//---------------------------------------------------------------------------------------------------------------
//
//  HAUD 2026.10.20
//
//
//  fb_DistributorByTicket
//  - uses 1 XtsStation via _ItfProcessCollector
//  - this instance checks its process list for an entry (Count > 0)
//      - pops ticket data from top of the list (GetHead)
//      - sends the mover to target stations according to bitmask in ST_PROCESS_DATA.wTarget
//
//  - inherits fb_Instance, which provides a design pattern in order to build different specific processes in a structured way
//  - used for targeting movers to predetermined bitmask of substations (one to many)
//
//
//  - constructed with fb_Instance main state (_eState) in addition to a substate (_eStateProgress)
//  - substate enables to handle procedures within main state by preventing race conditions 
//    with the help of small steps and decisions with clear separation from each other 
//
//---------------------------------------------------------------------------------------------------------------//
// This SOFTWARE is provided as an Exemple by THE PROVIDER "as is" and "with all faults." THE PROVIDER makes no  //
// representations or warranties of any kind concerning the safety, suitability, lack of viruses, inaccuracies,  //
// typographical errors, or other harmful components of this SOFTWARE. There are inherent dangers in the use of  //
// any software, and you are solely responsible for determining whether this SOFTWARE is compatible with your    //
// equipment and other software installed on your equipment. You are also solely responsible for the protection  //
// of your equipment and backup of your data, and THE PROVIDER will not be liable for any damages you may suffer //
// in connection with using, modifying, or distributing this SOFTWARE.                                           //
//---------------------------------------------------------------------------------------------------------------//
FUNCTION_BLOCK fb_DistributorByTicket EXTENDS fb_Instance
VAR
  //----------------------------------------------------------------------------------
  // outfeed target must be initialized with a valid target
  // I just use the default target that I am going to use in the basic process setup
  // this target is then updated and checked on arrival of a process ticket
  //----------------------------------------------------------------------------------
  _nProcessTarget               : E_INSTANCE;     // to whom am I connected --> to the data from the ticket
  //----------------------------------------------------------------------------------

  // target XTS station range
  _nTargetStationLast           : UINT;           // where does the target process end
  _nTargetStationFirst          : UINT;           // where does the target process start

  _WriteResult                  : ST_PROCESS_LIST_RESULT;   // last job written to target
  _DeleteResult                 : ST_PROCESS_LIST_RESULT;   // last job executed

  _nPrc                         : E_INSTANCE;
  _nTarget                      : E_INSTANCE;

  _idx                          : UINT;
  _nTargetIndex                 : ARRAY[1..SIZEOF(T_PROCESS)*8] OF USINT;

  _MoverInfo                    : ST_MOVER_INFO;      // Information from the Mover in Station
  _StationState                 : ST_STATION_STATE;   // BufferInfeed has only one XtsStation to work
END_VAR

//-----------------------------------------------------------------------------
//-----------------------------------------------------------------------------
// check pointer and interface
// connect Ctrl/State to _ItfProcessCollector
// set message device identification
//-----------------------------------------------------------------------------
IF NOT Check() THEN 
  RETURN; 
END_IF
//-----------------------------------------------------------------------------
// check command
//-----------------------------------------------------------------------------
_eCmd                                         := _stInstanceCtrl[_nProcess].Cmd;
IF (_eCmd <> _eCmdOld)
THEN
  CASE _eCmd
  OF
    E_INSTANCE_CMD.INIT:
      // clear init info
      _eInit                                  := _ItfProcessCollector[_nProcess].Init(FALSE);
  
      IF _ItfProcessList[_nProcess].InitList()  // clear linked list
      THEN
        Clear();
        _eStateInstance                       := E_INSTANCE_STATE.INIT;
        _eStateProgress                       := E_PROGRESS.PROGRESS_INIT;
      END_IF
  END_CASE
  CmdLog();
  _eCmdOld                                    := _eCmd;
END_IF
//-----------------------------------------------------------------------------
// cyclic information of mover and station
//-----------------------------------------------------------------------------
_StationState                                 := _ItfProcessCollector[_nProcess].GetStationState  (_ItfProcessCollector[_nProcess].StationLast);
//-----------------------------------------------------------------------------
//-----------------------------------------------------------------------------
// state machine for BufferInfeed work
//-----------------------------------------------------------------------------
CASE _eStateInstance
OF
  E_INSTANCE_STATE.NULL:
    // first cycle startup
    // initialize linked list, clears all entries
    IF _ItfProcessList[_nProcess].InitList()
    THEN
      _eInit                                  := _ItfProcessCollector[_nProcess].Init(FALSE);
      _eStateProgress                         := E_PROGRESS.PROGRESS_INIT;
      _eStateInstance                         := E_INSTANCE_STATE.INIT;
    END_IF


  E_INSTANCE_STATE.INIT:
    //-------------------------------------------------------------------------
    CASE _eStateProgress
    OF
    // E_INSTANCE_STATE.INIT:
    //-------------------------------------------------------------------------
      E_PROGRESS.PROGRESS_ERROR:
        IF (_nProcessTarget > 0) AND
           (_nProcessTarget < E_INSTANCE.INSTANCE_MAX)
        THEN
          _eStateProgress                     := E_PROGRESS.PROGRESS_INIT;
        END_IF

    // E_INSTANCE_STATE.INIT:
    //-------------------------------------------------------------------------
      E_PROGRESS.PROGRESS_INIT:
        IF NOT (_nProcessTarget > 0) OR
           NOT (_nProcessTarget < E_INSTANCE.INSTANCE_MAX)
        THEN
          _eStateProgress                     := E_PROGRESS.PROGRESS_ERROR;

        ELSE
          _eStateProgress                     := E_PROGRESS.PROGRESS_BUSY;
        END_IF

    // E_INSTANCE_STATE.INIT:
    //-------------------------------------------------------------------------
      E_PROGRESS.PROGRESS_BUSY:
        // wait for process collector check to be done
        //  - checks range of XtsStations
        //  - checks count of XtsStations
        IF (_stCollectorState.Check = E_PROCESS_CHECK.CHECK_DONE)
        THEN
          _eInit                              := _ItfProcessCollector[_nProcess].Init(TRUE);
  
          IF (_eInit = E_PROGRESS.PROGRESS_DONE)
          THEN
            IF NOT (_nProcessTarget > 0) OR
               NOT (_nProcessTarget < E_INSTANCE.INSTANCE_MAX)
            THEN
              // an invalid target you must have not
              _eStateProgress                 := E_PROGRESS.PROGRESS_ERROR;

              _stMsg.eType                    := E_MessageType.eMessageError;
              _stMsg.eSubdevice               := e_Subdevice.Instance_DistributorByTicket;
              _stMsg.iErrorNumber             := _nProcessTarget;
              _stMsg.sText                    := concat(TO_STRING(_eStateInstance), ': ProcessTarget: ');
              _stMsg.sText                    := concat(_stMsg.sText, TO_STRING(_eStateProgress));
              f_MessageSet(_stMsg);

            ELSE
              _ItfProcessCollector[_nProcess].Init(FALSE); // clear init procedure

              // initialization of BufferInfeed: _ItfProcessCollector with XtsStation
              _stCollectorCtrl.Cmd            := E_PROCESS_CTRL.PROCESS_DISABLE;  // switch off _ItfProcessCollector and XtsStation
              _eStateProgress                 := E_PROGRESS.PROGRESS_INIT;        // clear sub state
              _eStateInstance                 := E_INSTANCE_STATE.DISABLED;       // switch to disabled as default after startup
            END_IF
          END_IF
        END_IF
    END_CASE
END_CASE
//-----------------------------------------------------------------------------
// DISABLED:
//  - clear local list result data
//  - wait for enable from the outside
//-----------------------------------------------------------------------------
CASE _eStateInstance
OF
  E_INSTANCE_STATE.DISABLED:
    //-------------------------------------------------------------------------
    CASE _eStateProgress
    OF
      E_PROGRESS.PROGRESS_INIT:
        _stCollectorCtrl.Cmd                  := E_PROCESS_CTRL.PROCESS_DISABLE;  // switch off _ItfProcessCollector and XtsStation
        _eStateProgress                       := E_PROGRESS.PROGRESS_BUSY;
        // clear data for a new round
        memset(ADR(_stListResult), 0, SIZEOF(_stListResult));

        _stCollectorCtrl.ActivateStation      := 0; // clear activation mask of my process
        _stCollectorCtrl.NestMask             := 1; // my process target has one nest

        _nPrc                                 := _nProcess;
        _nTarget                              := _nProcessTarget;
    END_CASE
    // E_INSTANCE_STATE.DISABLED:
    //-------------------------------------------------------------------------
    CASE _eStateProgress
    OF
      E_PROGRESS.PROGRESS_BUSY:
        CASE _eCmd
        OF
          E_INSTANCE_CMD.ENABLE:              // turn it on!!
            _nPrc                             := _nProcess;
            _nTarget                          := _nProcessTarget;

            _eStateInstance                   := E_INSTANCE_STATE.DETECTION;
            _eStateProgress                   := E_PROGRESS.PROGRESS_BUSY;
  
            IF (_MessageLevel > E_MessageType.eMessageInfo)
            THEN
              _stMsg.eType                    := E_MessageType.eMessageVerbose;
              _stMsg.eSubdevice               := e_Subdevice.Instance_DistributorByTicket;
              _stMsg.iErrorNumber             := 0;
              _stMsg.sText                    := concat(TO_STRING(_eStateInstance), ': ');
              _stMsg.sText                    := concat(_stMsg.sText, TO_STRING(_eStateProgress));
              f_MessageSet(_stMsg);
            END_IF

        END_CASE
    END_CASE
END_CASE
//-----------------------------------------------------------------------------
// DETECTION: 
//  - check inked list and GetHead()
//  - copy job data
//  - switch on process
//-----------------------------------------------------------------------------
CASE _eStateInstance
OF
  E_INSTANCE_STATE.DETECTION:
    //-------------------------------------------------------------------------
    CASE _eStateProgress
    OF
      E_PROGRESS.PROGRESS_BUSY:
        IF (_eCmd = E_INSTANCE_CMD.DISABLE)
        THEN
          _eStateInstance                     := E_INSTANCE_STATE.DISABLED;
          _eStateProgress                     := E_PROGRESS.PROGRESS_INIT;

        ELSIF (_ItfProcessList[_nPrc].Count > 0)
        THEN
          // get new job order for my process
          // check my list for a new round of movers
          _stListResult                       := _ItfProcessList[_nPrc].GetHead();  // the list results carries information about the requirements of the target process (who and where)

          IF (_stListResult.wState <> 0)
          THEN
            // error in list results must not appear
            // if you land here, there is somethng wrong with the initialization or configuration of the linked list
            _eStateProgress                   := E_PROGRESS.PROGRESS_ERROR;

            _stMsg.eType                      := E_MessageType.eMessageError;
            _stMsg.eSubdevice                 := e_Subdevice.Process_LinkedList_GetHead;
            _stMsg.iErrorNumber               := _stListResult.wState;
            _stMsg.sText                      := concat(TO_STRING(_eStateInstance), ': _ListResult.wState: ');
            _stMsg.sText                      := concat(_stMsg.sText, TO_STRING(_eStateProgress));
            f_MessageSet(_stMsg);

          ELSE
            IF (_MessageLevel > E_MessageType.eMessageError)
            THEN
              _stMsg.eType                    := E_MessageType.eMessageInfo;
              _stMsg.eSubdevice               := e_Subdevice.Process_LinkedList_GetHead;
              _stMsg.iErrorNumber             := _nPrc;
              _stMsg.sText                    := concat(TO_STRING(_eStateInstance), ': ');
              _stMsg.sText                    := concat(_stMsg.sText, '_ListResult.stData.wTarget: ');
              _stMsg.sText                    := concat(_stMsg.sText, _ItfProcessCollector[_nPrc].BitsToString(_stListResult.stData.wTarget));
              f_MessageSet(_stMsg);
            END_IF

            _stProcessData                    := _stListResult.stData;  // list result contains data for target process

            IF (_stProcessData.wTarget > 0)
            THEN
              _eStateProgress                 := E_PROGRESS.PROGRESS_CHECK;

              IF (_MessageLevel = E_MessageType.eMessageBatch)
              THEN
                _stMsg.eType                  := E_MessageType.eMessageBatch;
                _stMsg.eSubdevice             := e_Subdevice.Instance_DistributorByTicket;
                _stMsg.iErrorNumber           := _nPrc;
                _stMsg.sText                  := concat(TO_STRING(_eStateProgress), ': ');
                _stMsg.sText                  := concat(_stMsg.sText, TO_STRING(e_message_batch.MSG_BATCH_JOB_STARTED));
                f_MessageSet(_stMsg);
              END_IF
            ELSE
              _DeleteResult                   := _ItfProcessList[_nPrc].RemoveHeadValue();
            END_IF

            // check target mask for entries
            IF NOT (_stProcessData.wTarget > 0)
            THEN
              _stMsg.eType                    := E_MessageType.eMessageWarning;
              _stMsg.eSubdevice               := e_Subdevice.Instance_DistributorByTicket;
              _stMsg.iErrorNumber             := 666;
              _stMsg.sText                    := concat(TO_STRING(_eStateInstance), ': ');
              _stMsg.sText                    := concat(_stMsg.sText, '_ProcessData.wTarget: ');
              _stMsg.sText                    := concat(_stMsg.sText, _ItfProcessCollector[_nProcess].BitsToString(_stProcessData.wTarget));
              f_MessageSet(_stMsg);
            END_IF
          END_IF
        END_IF
    END_CASE
    // E_INSTANCE_STATE.DETECTION
    //-------------------------------------------------------------------------
    CASE _eStateProgress
    OF
      E_PROGRESS.PROGRESS_CHECK:
        // do some plausibility checks on the ticket data
        IF NOT (_stProcessData.nTargetId > 0) OR
           NOT (_stProcessData.nTargetId < E_INSTANCE.INSTANCE_MAX) OR
           NOT (_stProcessData.nTargetId <> _nProcess)
        THEN
          _stMsg.eType                        := E_MessageType.eMessageError;
          _stMsg.eSubdevice                   := e_Subdevice.Instance_DistributorByTicket;
          _stMsg.iErrorNumber                 := _stProcessData.nTargetId;
          _stMsg.sText                        := concat(TO_STRING(_eStateInstance), ': _stProcessData.nTargetId: ');
          _stMsg.sText                        := concat(_stMsg.sText, TO_STRING(E_PROGRESS.PROGRESS_ERROR));
          f_MessageSet(_stMsg);

          // not a plausible target, delete ticket and go back to checking the list
          _DeleteResult                       := _ItfProcessList[_nPrc].RemoveHeadValue();
          _eStateProgress                     := E_PROGRESS.PROGRESS_BUSY;
        ELSE
          // update target data with ticket data
          _nTarget                            := _stProcessData.nTargetId;
          _nTargetStationLast                 := _ItfProcessCollector[_nTarget].StationLast;
          _nTargetStationFirst                := _ItfProcessCollector[_nTarget].StationFirst;

          IF (_ItfProcessCollector[_nTarget].ProcessState.Check = E_PROCESS_CHECK.CHECK_DONE)
          THEN
            _eStateProgress                   := E_PROGRESS.PROGRESS_WORKING;

            IF (_MessageLevel > E_MessageType.eMessageWarning)
            THEN
              _stMsg.eType                    := E_MessageType.eMessageInfo;
              _stMsg.eSubdevice               := e_Subdevice.Instance_DistributorByTicket;
              _stMsg.iErrorNumber             := _stProcessData.nTargetId;
              _stMsg.sText                    := concat(TO_STRING(_stProcessData.nProcessId), ': _stProcessData.nTargetId: ');
              _stMsg.sText                    := concat(_stMsg.sText, TO_STRING(_eStateProgress));
              f_MessageSet(_stMsg);
            END_IF
          END_IF
        END_IF
    END_CASE
    // E_INSTANCE_STATE.DETECTION
    //-------------------------------------------------------------------------
    CASE _eStateProgress
    OF
      E_PROGRESS.PROGRESS_WORKING:
        // check for disabled process interface state
        CASE _stCollectorState.State
        OF
          E_PROCESS_STATE.PROCESS_DISABLE:

          CASE _stCollectorState.Result
          OF
            E_PROGRESS.PROGRESS_BUSY:         // busy from _State.Result means, waiting for input
              // now the preparation for the target process may begin
              _stCollectorCtrl.Cmd               := E_PROCESS_CTRL.PROCESS_ENABLE; // switch on my state machine in _ItfProcessCollector
              _stCollectorCtrl.ActivateStation   := 1;                             // enable my XtsStation in _ItfProcessCollector (BufferInfeed has only one XtsStation)

              _eStateInstance                 := E_INSTANCE_STATE.ENABLED;         // go check if my process is switched on
              _eStateProgress                 := E_PROGRESS.PROGRESS_INIT;         // reset substate

              IF (_MessageLevel > E_MessageType.eMessageInfo)
              THEN
                _stMsg.eType                  := E_MessageType.eMessageVerbose;
                _stMsg.eSubdevice             := e_Subdevice.Instance_DistributorByTicket;
                _stMsg.iErrorNumber           := 0;
                _stMsg.sText                  := concat(TO_STRING(_eStateInstance), ': ');
                _stMsg.sText                  := concat(_stMsg.sText, TO_STRING(_eStateProgress));
                f_MessageSet(_stMsg);
              END_IF
          END_CASE
        END_CASE
    END_CASE
END_CASE
//-----------------------------------------------------------------------------
// ENABLED
//  - check process for enabled stations from list entry
//  - switch to sending
//  - allow movers to be sent
//-----------------------------------------------------------------------------
CASE _eStateInstance
OF
  E_INSTANCE_STATE.ENABLED:
    //-------------------------------------------------------------------------
    CASE _eStateProgress
    OF
      E_PROGRESS.PROGRESS_INIT:
        CASE _stCollectorState.State
        OF
          E_PROCESS_STATE.PROCESS_ENABLE:
          CASE _stCollectorState.Result
          OF
            E_PROGRESS.PROGRESS_BUSY:
              // now my process and all XtsStations within are switched on
              // check infeed into my process
              _stCollectorCtrl.Cmd            := E_PROCESS_CTRL.PROCESS_STATIONS_SEND; // tells my process to go check the infeed
              _eStateProgress                 := E_PROGRESS.PROGRESS_BUSY; // go check how the infeed into my process is doing

              IF (_MessageLevel > E_MessageType.eMessageWarning)
              THEN
                _stMsg.eType                  := E_MessageType.eMessageInfo;
                _stMsg.eSubdevice             := e_Subdevice.Instance_DistributorByTicket;
                _stMsg.iErrorNumber           := _StationState.nMoverId;
                _stMsg.sText                  := concat(TO_STRING(_eStateInstance), ': ');
                _stMsg.sText                  := concat(_stMsg.sText, TO_STRING(_eStateProgress));
                f_MessageSet(_stMsg);
              END_IF
          END_CASE
        END_CASE
    END_CASE
    // E_INSTANCE_STATE.ENABLED:
    //-------------------------------------------------------------------------
    CASE _eStateProgress
    OF
      E_PROGRESS.PROGRESS_BUSY:
        CASE _stCollectorState.State
        OF
          E_PROCESS_STATE.PROCESS_STATIONS_OUTFEED:
          CASE _stCollectorState.Result       // if collector is ready to send mover
          OF
            E_PROGRESS.PROGRESS_BUSY:
              // check if the mover is in range
              IF (_rCheckPositionEnd > _rCheckPositionStart)
              THEN
                IF (_StationState.rMoverModPos > _rCheckPositionStart) AND
                   (_StationState.rMoverModPos < _rCheckPositionEnd)
                THEN
                  _eStateProgress             := E_PROGRESS.PROGRESS_PREPARE;
                END_IF
              ELSE
                IF (_StationState.rMoverModPos > _rCheckPositionStart) OR
                   (_StationState.rMoverModPos < _rCheckPositionEnd)
                THEN
                  _eStateProgress             := E_PROGRESS.PROGRESS_PREPARE;
                END_IF
              END_IF
          END_CASE
        END_CASE
    END_CASE
    // E_INSTANCE_STATE.ENABLED:
    //-------------------------------------------------------------------------
    CASE _eStateProgress
    OF
      E_PROGRESS.PROGRESS_PREPARE:
        // now we know the mover is in range
        // continue to finish
        _stCollectorCtrl.Cmd                  := E_PROCESS_CTRL.PROCESS_STATIONS_SEND;

        _eStateInstance                       := E_INSTANCE_STATE.FINISH;   // go get data ready for outfeed
        _eStateProgress                       := E_PROGRESS.PROGRESS_INIT;  // reset substate

        IF (_MessageLevel > E_MessageType.eMessageError)
        THEN
          _stMsg.eType                        := E_MessageType.eMessageInfo;
          _stMsg.eSubdevice                   := e_Subdevice.Instance_DistributorByTicket;
          _stMsg.iErrorNumber                 := _StationState.nMoverId;
          _stMsg.sText                        := concat(TO_STRING(_eStateInstance), ': ');
          _stMsg.sText                        := concat(_stMsg.sText, TO_STRING(_eStateProgress));
          f_MessageSet(_stMsg);
        END_IF
    END_CASE
END_CASE
//-----------------------------------------------------------------------------
// FINISH:
//  - write target (Last to First)
//  - delete target bit from linked list result (_ProcessData.wTarget)
//  - send out mover
//  - check _ProcessData.wTarget for next mover
//  - check if all movers in job were sent (ProcessData.wTarget = 0)
//  - RemoveHead() from my list
//  - AddTail() at TargetProcess
//  - check to proceed
//-----------------------------------------------------------------------------
CASE _eStateInstance
OF
  E_INSTANCE_STATE.FINISH:
    //-------------------------------------------------------------------------
    CASE _eStateProgress
    OF
      E_PROGRESS.PROGRESS_INIT:
      // check bit mask for sending mover to required targets
      // get target index for mover from process list entry
      FOR _idx := _nTargetStationLast TO _nTargetStationFirst BY(-1)
      DO
        IF (ItfProcessCollector[_nPrc].BitGet(_stProcessData.wTarget, _idx-_nTargetStationFirst))
        THEN
          _eStateProgress                     := E_PROGRESS.PROGRESS_BUSY;

          _nTargetIndex[1]                    := TO_USINT(_idx);
          _ItfProcessCollector[_nPrc].TargetIndex := _nTargetIndex; // write Xts target onto my ProcessCollector interface

          // got the target, now delete the just found bit of this job
          _stProcessData.wTarget              := _ItfProcessCollector[_nPrc].
                                                 BitDel(_stProcessData.wTarget, _idx-_nTargetStationFirst);

          IF (_MessageLevel > E_MessageType.eMessageVerbose)
          THEN
            _stMsg.eType                      := E_MessageType.eMessageSentient;
            _stMsg.eSubdevice                 := e_Subdevice.Instance_DistributorByTicket;
            _stMsg.iErrorNumber               := _idx;
            _stMsg.sText                      := concat('_ProcessData.wTarget: ', 
                                                 _ItfProcessCollector[_nPrc].BitsToString(_stProcessData.wTarget));
            f_MessageSet(_stMsg);
          END_IF
          EXIT;
        END_IF
      END_FOR
    END_CASE
    // E_INSTANCE_STATE.FINISH:
    //-------------------------------------------------------------------------
    CASE _eStateProgress
    OF
      E_PROGRESS.PROGRESS_BUSY:
        CASE _stCollectorState.State
        OF
          E_PROCESS_STATE.PROCESS_STATIONS_OUTFEED: // double check my process' state
          CASE _stCollectorState.Result
          OF
            E_PROGRESS.PROGRESS_BUSY:
              // now data is prepared and copied to the right places
              _stCollectorCtrl.Cmd            := E_PROCESS_CTRL.PROCESS_STATIONS_OUTFEED; // tell my process to release the mover
              _eStateProgress                 := E_PROGRESS.PROGRESS_CHECK; // go check for more to do

              IF (_MessageLevel > E_MessageType.eMessageInfo)
              THEN
                _stMsg.eType                  := E_MessageType.eMessageVerbose;
                _stMsg.eSubdevice             := e_Subdevice.Instance_DistributorByTicket;
                _stMsg.iErrorNumber           := _nPrc;
                _stMsg.sText                  := concat(TO_STRING(_eStateInstance), ': ');
                _stMsg.sText                  := concat(_stMsg.sText, TO_STRING(_eStateProgress));
                f_MessageSet(_stMsg);
              END_IF
          END_CASE
        END_CASE
    END_CASE
    // E_INSTANCE_STATE.FINISH:
    //-------------------------------------------------------------------------
    CASE _eStateProgress
    OF
      E_PROGRESS.PROGRESS_CHECK:
        CASE _stCollectorState.State
        OF
          E_PROCESS_STATE.PROCESS_DISABLE:
            IF (_stProcessData.wTarget <> 0)
            THEN
              _stCollectorCtrl.Cmd               := E_PROCESS_CTRL.PROCESS_ENABLE; // switch on my state machine in _ItfProcessCollector
              _stCollectorCtrl.ActivateStation   := 1;                             // enable my XtsStation in _ItfProcessCollector (BufferInfeed has only one XtsStation)

              _eStateInstance                 := E_INSTANCE_STATE.ENABLED;         // go check if my process is switched on
              _eStateProgress                 := E_PROGRESS.PROGRESS_INIT;         // reset substate

              IF (_MessageLevel > E_MessageType.eMessageInfo)
              THEN
                _stMsg.eType                  := E_MessageType.eMessageVerbose;
                _stMsg.eSubdevice             := e_Subdevice.Instance_DistributorByTicket;
                _stMsg.iErrorNumber           := _nPrc;
                _stMsg.sText                  := concat(TO_STRING(_eStateInstance), ': ');
                _stMsg.sText                  := concat(_stMsg.sText, TO_STRING(_eStateProgress));
                f_MessageSet(_stMsg);
              END_IF
            ELSE
              // job done, all movers were sent
              // job done, delete from top of my list
              _DeleteResult                   := _ItfProcessList[_nPrc].RemoveHeadValue();

              IF (_DeleteResult.wState <> 0)
              THEN
                // deleting from list must be successful
                // IF you land here, there is something wrong with initialization or configuration of the linked list
                _eStateProgress               := E_PROGRESS.PROGRESS_ERROR;
              ELSE
                _eStateProgress               := E_PROGRESS.PROGRESS_WORKING; // job is done, now go and write ticket to _nTargetProcess
              END_IF
            END_IF 
        END_CASE
    END_CASE
    // E_INSTANCE_STATE.FINISH:
    //-------------------------------------------------------------------------
    CASE _eStateProgress
    OF
      E_PROGRESS.PROGRESS_WORKING:
        // write process ticket, then go back up
        //_WriteResult                          := _ItfProcessList[_nTarget].AddTailValue(_stListResult.stData);

        IF (_WriteResult.wState <> 0)
        THEN
          // adding to target list must be successful on the first try
          // IF you land here, there is something wrong with initialization or configuration of the linked list
          _eStateProgress                     := E_PROGRESS.PROGRESS_ERROR;
        ELSE
          _eStateProgress                     := E_PROGRESS.PROGRESS_DONE;

          IF (_MessageLevel > E_MessageType.eMessageError)
          THEN
            _stMsg.eType                      := E_MessageType.eMessageInfo;
            _stMsg.eSubdevice                 := e_Subdevice.Process_LinkedList_AddTail;
            _stMsg.iErrorNumber               := _nTarget;
            _stMsg.sText                      := concat(TO_STRING(_eStateInstance), ': ');
            _stMsg.sText                      := concat(_stMsg.sText, TO_STRING(_eStateProgress));
            //f_MessageSet(_stMsg);
          END_IF
          IF (_MessageLevel = E_MessageType.eMessageBatch)
          THEN
            _stMsg.eType                      := E_MessageType.eMessageBatch;
            _stMsg.eSubdevice                 := e_Subdevice.Instance_DistributorByTicket;
            _stMsg.iErrorNumber               := _nPrc;
            _stMsg.sText                      := concat(TO_STRING(_eStateProgress), ': ');
            _stMsg.sText                      := concat(_stMsg.sText, TO_STRING(e_message_batch.MSG_BATCH_JOB_DONE));
            f_MessageSet(_stMsg);
          END_IF
        END_IF
    END_CASE
    // E_INSTANCE_STATE.FINISH:
    //-------------------------------------------------------------------------
    CASE _eStateProgress
    OF
      E_PROGRESS.PROGRESS_DONE:
        //----------------------------------
        //  wait for command from higher up
        //----------------------------------
        CASE _eCmd
        OF
          // command to disable required
          E_INSTANCE_CMD.DISABLE:
            _eStateInstance                   := E_INSTANCE_STATE.DISABLED;
            _eStateProgress                   := E_PROGRESS.PROGRESS_INIT;

            IF (_MessageLevel > E_MessageType.eMessageInfo)
            THEN
              _stMsg.eType                    := E_MessageType.eMessageVerbose;
              _stMsg.eSubdevice               := e_Subdevice.Instance_DistributorByTicket;
              _stMsg.iErrorNumber             := _nPrc;
              _stMsg.sText                    := concat(TO_STRING(_eStateInstance), ': ');
              _stMsg.sText                    := concat(_stMsg.sText, TO_STRING(_eStateProgress));
              f_MessageSet(_stMsg);
            END_IF
        END_CASE
    END_CASE
END_CASE
//-----------------------------------------------------------------------------
//-----------------------------------------------------------------------------
_stInstanceState[_nProcess].ProcessIdentity   := _nProcess;
_stInstanceState[_nProcess].ProcessState      := _eStateInstance;
_stInstanceState[_nProcess].ProcessProgress   := _eStateProgress;
//-----------------------------------------------------------------------------
//-----------------------------------------------------------------------------
_stInstanceState[_nProcess].CollectorState    := _stCollectorState.State;
_stInstanceState[_nProcess].CollectorProgress := _stCollectorState.Result;
_stInstanceState[_nProcess].CollectorCheck    := _stCollectorState.Check;
_stInstanceState[_nProcess].StationCount      := _ItfProcessCollector[_nProcess].StationCount;
_stInstanceState[_nProcess].QueueProcessCount := _ItfProcessCollector[_nProcess].QueueProcessCount;
_stInstanceState[_nProcess].ListCount         := TO_UINT(_ItfProcessList[_nProcess].Count);
//-----------------------------------------------------------------------------
//-----------------------------------------------------------------------------

METHOD Clear : BOOL
VAR_INPUT
END_VAR
memset(ADR(_nTargetIndex), 0, SIZEOF(_nTargetIndex));

//_eStateInstance                         := E_INSTANCE_STATE.DISABLED;
_eStateProgress                 := E_PROGRESS.PROGRESS_INIT;

Clear                           := TRUE;
END_METHOD

PROPERTY ProcessTarget : E_INSTANCE
GET
ProcessTarget := _nProcessTarget;
END_GET
SET
_nProcessTarget := ProcessTarget;
END_SET
END_PROPERTY

END_FUNCTION_BLOCK

(* stored: Version 1.1.0.1
   POU fb_DistributorByTicket: Id {e80657f1-fb68-402a-bc07-d7a99c278aae}, SpecialFunc None
   Method Clear: Id {1b71cdc4-bfaa-46a0-b309-fc130d1116e3}
   Property ProcessTarget: Id {6107843f-d643-4898-8d2d-3433ca504ba7}
   Get Get: Id {f141dcd0-3a08-4969-8e39-8d8a4c21d219}
   Set Set: Id {b5bb18f1-16f9-4669-9e34-58d2035ce8c2} *)
